// TIA Portal V20 export
// export: Created 2026-10-12T04:58:22.6426041Z, ExportSetting WithDefaults, DisplayName Totally Integrated Automation Portal, DisplayVersion V20, DisplayName TIA Portal Openness, DisplayVersion V20, DisplayName TIA Portal Teamcenter Gateway, DisplayVersion V20, DisplayName TIA Portal Version Control Interface, DisplayVersion V20, DisplayName SINAMICS Startdrive Advanced, DisplayVersion V20 SP1 Update 2, DisplayName SINAMICS Startdrive G110M, G120, G120C, G120D, G120P, G115D, DisplayVersion V20 SP1 Update 2, DisplayName SINAMICS Startdrive G130, G150, S120, S150, SINAMICS MV, G220, S200, S210, DisplayVersion V20 SP1 Update 2, DisplayName STEP 7 Professional, DisplayVersion V20, DisplayName STEP 7 Safety, DisplayVersion V20, DisplayName WinCC Basic/Comfort/Advanced, DisplayVersion V20, DisplayName WinCC Professional, DisplayVersion V20, DisplayName WinCC Unified, DisplayVersion V20
FUNCTION "FRK_CfgDef_DeclarationCylinder" : Void   // FC123, SCL
{ S7_Optimized_Access := 'TRUE' }
VERSION : 0.1
// stored: AutoNumber true, IsIECCheckEnabled false, SetENOAutomatically false, UDAEnableTagReadback false
   VAR_INPUT
      FieldIndex : Int;
   END_VAR
BEGIN

   "FRK_ConfigScratch".Entry := "FRK_ConfigScratch".Blank;
   CASE #FieldIndex OF
       1:
           "FRK_ConfigScratch".Entry.WriteKey := 'timeout';
           "FRK_ConfigScratch".Entry.WriteRevision := UDINT#1;
           "FRK_ConfigScratch".Entry.Item := WSTRING#'ParCfg/Timeout';
           "FRK_ConfigScratch".Entry.ConfigKind := 0;
           "FRK_ConfigScratch".Entry.ValueType := 3;
           "FRK_ConfigScratch".Entry.Writable := TRUE;
           "FRK_ConfigScratch".Entry.RequiresReady := TRUE;
           "FRK_ConfigScratch".Entry.HasMinimum := TRUE;
           "FRK_ConfigScratch".Entry.HasMaximum := TRUE;
           "FRK_ConfigScratch".Entry.Minimum := 1.0;
           "FRK_ConfigScratch".Entry.Maximum := 60000.0;
           "FRK_ConfigScratch".Entry.LabelKey := 'test.config.timeout';
           "FRK_ConfigScratch".Storage := 7;
           "FRK_ConfigScratch".Schema := 4;
           "FRK_ConfigScratch".Minimum := 1.0;
           "FRK_ConfigScratch".Maximum := 60000.0;
           "FRK_ConfigScratch".MaxLength := 0;
           "FRK_ConfigScratch".MinRead := 0;
           "FRK_ConfigScratch".MinWrite := 0;
       2:
           "FRK_ConfigScratch".Entry.WriteKey := 'preset';
           "FRK_ConfigScratch".Entry.WriteRevision := UDINT#2;
           "FRK_ConfigScratch".Entry.Item := WSTRING#'ParCfg/Preset';
           "FRK_ConfigScratch".Entry.ConfigKind := 0;
           "FRK_ConfigScratch".Entry.ValueType := 0;
           "FRK_ConfigScratch".Entry.Writable := TRUE;
           "FRK_ConfigScratch".Entry.RequiresReady := TRUE;
           "FRK_ConfigScratch".Entry.HasMinimum := TRUE;
           "FRK_ConfigScratch".Entry.HasMaximum := TRUE;
           "FRK_ConfigScratch".Entry.Minimum := 0.0;
           "FRK_ConfigScratch".Entry.Maximum := 1000.0;
           "FRK_ConfigScratch".Entry.LabelKey := 'test.config.preset';
           "FRK_ConfigScratch".Storage := 3;
           "FRK_ConfigScratch".Schema := 4;
           "FRK_ConfigScratch".Minimum := 0.0;
           "FRK_ConfigScratch".Maximum := 1000.0;
           "FRK_ConfigScratch".MaxLength := 0;
           "FRK_ConfigScratch".MinRead := 0;
           "FRK_ConfigScratch".MinWrite := 1;
       ELSE
           RETURN;
   END_CASE;
END_FUNCTION
